// TIA Portal project "Types" (V21)

(* hardware
DEVICE "PLC_Types"  S7-1500 station
   slot 0: "Rail_0"  Rack  6ES7 590-1***0-0AA0
   slot 1: "PLC_Types"  CPU 1516-3 PN/DP  6ES7 516-3AN02-0AB0  V2.9
      slot 3: "CPU display_1"  6ES7591-1BA00-0AA0
      slot 32768: "PROFINET interface_1"  X1
         slot 32769: "Port_1"  X1 P1
         slot 32770: "Port_2"  X1 P2
      slot 33024: "PROFINET interface_2"  X2
         slot 33025: "Port_1"  X2 P1
      slot 33280: "DP interface_1"  X3
      slot 34817: "Virtual CP interface port_1"  Virtual CP interface port  Virtual CP interface port
*)

// ===== PLC "PLC_Types"  CPU 1516-3 PN/DP =====

TYPE "typeInner"
   STRUCT
      flag : Bool := TRUE;   // A flag with a start value
      count : Int := 7;   // A counter with a start value
      value : Real := 2.5;   // A value with a start value
   END_STRUCT;
END_TYPE

TYPE "typeOuter"
   STRUCT
      inner : "typeInner";   // One inner type
      list : Array[1..3] of "typeInner";   // Three of them
      matrix : Array[0..1, 0..2] of Int;   // Two dimensions
      nested : Struct   // A struct in a struct
         "a" : Bool := TRUE;
         "b" : Struct
            c : Real := 1.5;
            d : Array[0..1] of Bool;
         END_STRUCT;
      END_STRUCT;
      text : String[16] := 'outer';   // A short string
   END_STRUCT;
END_TYPE

DATA_BLOCK "AllTypes"   // DB1
TITLE = Every elementary type
{ S7_Optimized_Access := 'TRUE' }
VERSION : 0.1
   VAR
      aBool : Bool := TRUE;
      aByte : Byte := 16#AB;
      aWord : Word := 16#ABCD;
      aDWord : DWord := 16#DEAD_BEEF;
      aLWord : LWord := 16#0123_4567_89AB_CDEF;
      aSInt : SInt := -5;
      aUSInt : USInt := 200;
      aInt : Int := -1234;
      aUInt : UInt := 60000;
      aDInt : DInt := -100000;
      aUDInt : UDInt := 4_000_000_000;
      aLInt : LInt := -9_000_000_000;
      aULInt : ULInt := 18_000_000_000_000_000_000;
      aReal : Real := 3.25;
      aLReal : LReal := -1.0E-10;
      aTime : Time := T#1D_2H_3M_4S_5MS;
      aLTime : LTime := LT#1S_500NS;
      aS5Time : S5Time := S5T#10S;
      aDate : Date := D#2024-02-29;
      aTimeOfDay : Time_Of_Day := TOD#12:34:56.789;
      aLTimeOfDay : LTime_Of_Day := LTOD#12:34:56.123456789;
      aDateAndTime : Date_And_Time := DT#2024-02-29-12:00:00;
      anLDT : LDT := LDT#2024-02-29-12:00:00.123456789;
      aDTL : DTL := DTL#2024-02-29-12:00:00;
      aChar : Char := 'A';
      aWChar : WChar := WCHAR#'B';
      aString : String := 'hello';
      aShortString : String[10] := 'short';
      aWString : WString := WSTRING#'wide';
      anArray : Array[0..3] of Int;
      aMatrix : Array[1..2, 1..3] of Real;
      anArrayOfStruct : Array[1..2] of Struct
         on : Bool;
         speed : Int;
      END_STRUCT;
   END_VAR
BEGIN
   anArray[0] := 1;
   anArray[1] := 2;
   anArray[2] := 3;
   anArray[3] := 4;
   aMatrix[1,1] := 0.5;
   aMatrix[1,2] := 1.5;
   aMatrix[1,3] := 2.5;
   aMatrix[2,1] := 3.5;
   aMatrix[2,2] := 4.5;
   aMatrix[2,3] := 5.5;
   anArrayOfStruct[1].on := TRUE;
   anArrayOfStruct[2].on := TRUE;
   anArrayOfStruct[1].speed := 100;
   anArrayOfStruct[2].speed := 100;
END_DATA_BLOCK

DATA_BLOCK "Retained"   // DB2
{ S7_Optimized_Access := 'TRUE' }
VERSION : 0.1
   VAR RETAIN
      kept : DInt := 42;   // Survives a power cycle
      keptText : String[8] := 'kept';
   END_VAR
   VAR
      lost : DInt := 7;   // Starts again from its start value
   END_VAR
BEGIN
END_DATA_BLOCK

DATA_BLOCK "Classic"   // DB3
{ S7_Optimized_Access := 'FALSE' }
VERSION : 0.1
   VAR
      first : Bool := TRUE;   // At offset 0.0
      second : Int := 22;   // At offset 2.0
      third : Real := 3.0;   // At offset 4.0
      fourth : Array[1..4] of Byte;
   END_VAR
BEGIN
   fourth[1] := 16#0001;
   fourth[2] := 16#0002;
   fourth[3] := 16#0003;
   fourth[4] := 16#0004;
END_DATA_BLOCK

DATA_BLOCK "Settings"   // DB4
{ S7_Optimized_Access := 'TRUE' }
VERSION : 0.1
BEGIN
   inner.count := 11;
   list[2].value := 9.75;
   matrix[1,2] := 12;
   nested."b".c := -4.5;
   text := 'settings';
END_DATA_BLOCK

DATA_BLOCK "InterfaceData"   // DB5
{ S7_Optimized_Access := 'TRUE' }
VERSION : 0.1
// stored: InstanceOfName Interface
"Interface"
BEGIN
   setpoint := 75.0;
   state := 4;
END_DATA_BLOCK

FUNCTION_BLOCK "Interface"   // FB1, SCL
TITLE = Every section of an interface
{ S7_Optimized_Access := 'TRUE' }
VERSION : 0.1
// Inputs, outputs, in-outs, statics, temporaries and constants, with start values.
   VAR_INPUT
      enable : Bool := TRUE;   // Input with a start value
      setpoint : Real := 50.0;
      config : "typeInner";   // A data type as input
   END_VAR
   VAR_OUTPUT
      busy : Bool;
      result : DInt := -1;
   END_VAR
   VAR_IN_OUT
      shared : "typeOuter";   // A data type passed by reference
   END_VAR
   VAR
      state : Int := 3;
      history : Array[1..5] of Real;
      delay : TON_TIME;
      local : "typeInner";
   END_VAR
   VAR_TEMP
      scratch : DInt;
   END_VAR
   VAR CONSTANT
      LIMIT_HIGH : Real := 100.0;   // A constant
      STEPS : Int := 5;
      LABEL : String := 'iface';
   END_VAR
   // history[1] := 1.0;
   // history[2] := 2.0;
   // history[3] := 3.0;
   // history[4] := 4.0;
   // history[5] := 5.0;
BEGIN

    #delay(IN := #enable,
           PT := T#1S);
    #busy := #enable AND NOT #delay.Q;
    #scratch := #state * #STEPS;
    IF #setpoint > #LIMIT_HIGH THEN
        #result := -1;
    ELSE
        #result := #scratch + #shared.inner.count + #config.count;
    END_IF;
    #history[1] := #setpoint;
    #local := #config;
END_FUNCTION_BLOCK

FUNCTION "Average" : LReal   // FC1, SCL
TITLE = Average of an array
{ S7_Optimized_Access := 'TRUE' }
VERSION : 0.1
// A function with a return value, an array passed in, and temporary data.
   VAR_INPUT
      values : Array[0..9] of LReal;   // The values
      count : Int;   // How many of them count
   END_VAR
   VAR_TEMP
      sum : LReal;
      i : Int;
   END_VAR
BEGIN

    #sum := 0.0;
    FOR #i := 0 TO LIMIT(MN := 0, IN := #count, MX := 10) - 1 DO
        #sum := #sum + #values[#i];
    END_FOR;
    IF #count > 0 THEN
        #Average := #sum / INT_TO_LREAL(#count);
    ELSE
        #Average := 0.0;
    END_IF;
END_FUNCTION